SUBAPPLICATION AX_TO_QXA_Option (* Reiner physischer Ausgang: AX-Zustand auf logiBUS_QXA, aktiviert per AOption (INIT/QI ueber AOption_X_TO_EVENT, INIT_CNF echt von DigitalOutput.INITO). *)
  (* Standard: 61499-2; Description: Copyright (c) 2026 Meisterschulen am Ostbahnhof This program and the accompanying materials are made available under the terms of the Eclipse Public License 2.0 which is available at https://www.eclipse.org/legal/epl-2.0/ SPDX-License-Identifier: EPL-2.0 *)
  (* Version 1.0, 2026-10-17, Franz Höpfinger, Meisterschulen am Ostbahnhof, initial implementation - Ausgangs-Teil von AX_TO_QXA_BG_PUBLISH_SWITCHPIC_OPT als eigener Baustein (Franz: an AOption_T_2_Klassisch ein reiner OUT-Baustein), Muster wie OptionalGroup_001. *)
  PACKAGE MyLib::sys;
  IMPORT logiBUS::io::DQ::logiBUS_DO;
  IMPORT logiBUS::io::DQ::logiBUS_DO_S;
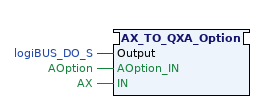
  VAR_INPUT
    Output : logiBUS::io::DQ::logiBUS_DO_S := logiBUS_DO::Invalid; (* Identify the Output Output_Q1..Q12 *)
  END_VAR
  SOCKETS
    AOption_IN : Option::AOption; (* Aktiviert/deaktiviert den Ausgang *)
    IN : adapter::types::unidirectional::AX; (* Fertiger AX-Zustand fuer den Ausgang *)
  END_SOCKETS
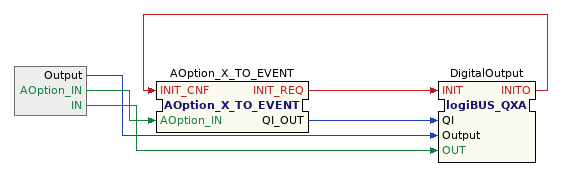
  FBS
    AOption_X_TO_EVENT : Option::conversion::AOption_X_TO_EVENT;
    DigitalOutput : logiBUS::io::DQ::logiBUS_QXA;
  END_FBS
  EVENT_CONNECTIONS
    AOption_X_TO_EVENT.INIT_REQ TO DigitalOutput.INIT;
    DigitalOutput.INITO TO AOption_X_TO_EVENT.INIT_CNF;
  END_CONNECTIONS
  DATA_CONNECTIONS
    AOption_X_TO_EVENT.QI_OUT TO DigitalOutput.QI;
    Output TO DigitalOutput.Output;
  END_CONNECTIONS
  ADAPTER_CONNECTIONS
    AOption_IN TO AOption_X_TO_EVENT.AOption_IN;
    IN TO DigitalOutput.OUT;
  END_CONNECTIONS
END_SUBAPPLICATION
